# EPICS substitutions: iocs/motor/ims-ioc/db/IM483.substitutions
# C's iocIms IM483.substitutions, P and C from st-im483sm.cmd.
file "$(MOTOR)/db/motor.db"
{
pattern
{N, M,       DTYP,      S, DESC,         EGU,     DIR, VELO, VBAS, ACCL, BDST, BVEL, BACC, MRES, PREC, DHLM, DLLM, INIT}
{1, "m$(N)", "IM483SM", 0, "motor $(N)", degrees, Pos, 1,    .1,   .2,   0,    1,    .2,   0.01, 5,    100,  -100, ""}
}
